// TIA Portal V20 export
Screen "5056 - G05 Pumps"  NonexNone, Number=5056
  ScreenLayer "Layer_0"
    FaceplateInstance "Faceplate_1"  FaceplateTypeName=_Library@$@Redesign@$@Faceplate@$@faceplatePump20Operate V 0.0.2
    FaceplateInstance "Faceplate_2"  FaceplateTypeName=_Library@$@Redesign@$@Faceplate@$@faceplateSafetyDevice V 1.0.0
    FaceplateInstance "Faceplate_3"  FaceplateTypeName=_Library@$@faceplateMissing V 0.1.0
